INTERFACE I_Conveyor EXTENDS I_Command, I_Status

END_INTERFACE

(* stored: Version 1.1.0.1, ProductVersion 3.1 *)
